FUNCTION_BLOCK Overpressure (* Basic Function Block Type *)
  (* Standard: 61499-2 *)
  (* Version 0.0, 6/22/2016, Andrei, nxtControl GmbH, Template *)
  PACKAGE Main;
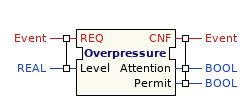
  EVENT_INPUT
    REQ WITH Level; (* Normal Execution Request *)
  END_EVENT
  EVENT_OUTPUT
    CNF WITH Attention, Permit; (* Execution Confirmation *)
  END_EVENT
  VAR_INPUT
    Level : REAL; (* Input event qualifier *)
  END_VAR
  VAR_OUTPUT
    Attention : BOOL; (* Output event qualifier *)
    Permit : BOOL := TRUE;
  END_VAR
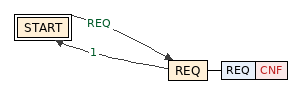
  EC_STATES
    START; (* Initial State *)
    REQ : REQ -> CNF;
  END_STATES
  EC_TRANSITIONS
    START TO REQ := REQ;
    REQ TO START := 1;
  END_TRANSITIONS
  ALGORITHM REQ IN ST: (* Initialization algorithm *)
IF Level >= 450.0 THEN
	Attention := TRUE;
ELSE
	Attention := FALSE;
END_IF;
IF Level > 599.0 THEN
	Permit := FALSE;
ELSE
	Permit := TRUE;
END_IF;
  END_ALGORITHM
END_FUNCTION_BLOCK
